// TIA Portal V21 export
FUNCTION_BLOCK "GuardSafety"   // FB4, F_FBD
{ S7_Optimized_Access := 'TRUE' }
// Main safety block of the guard's F-runtime group.
   VAR
      guard : "Guard";
      hornOn : Bool;
   END_VAR
BEGIN

REGION Network 1: Guard
   // The horn is on while the guard is open.
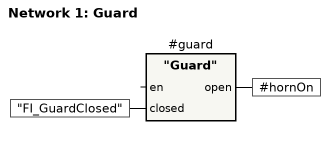
   #guard(closed := "FI_GuardClosed", open => #hornOn);   // "Guard"
END_REGION
END_FUNCTION_BLOCK
